Fanuc KAREL source: kc00039.KL

-- PROVISIONAL review KL for V940-1; original PC SHA256 a3de00926e4ed159da5d7aff602eb50377b7e1f1824aacf54da72a1891f8539a
-- Incomplete behavior may be omitted. Consult companion uncertainty JSON. Do not deploy.
PROGRAM KC00039
%NOLOCKGROUP
BEGIN
  -- V9_ZERO_TABLE_METADATA_HINT layout=0001; no indexed target words; source/name/runtime held
  -- UNRESOLVED_PC offsets 5-32; opcodes 27,22,22,1C,22,76
  -- UNRESOLVED_PC offsets 37-41; opcodes 7F
END KC00039
